// TIA Portal V21 export
// export: Created 2026-11-10T19:11:42.2574666Z, ExportSetting WithDefaults, DisplayName Totally Integrated Automation Portal, DisplayVersion V21 Update 3, DisplayName STEP 7 Professional, DisplayVersion V21 Update 3, DisplayName STEP 7 Safety, DisplayVersion V21, DisplayName Tech WebApplication, DisplayVersion V21, DisplayName WinCC Basic/Comfort/Advanced, DisplayVersion V21 Update 3, DisplayName WinCC Unified, DisplayVersion V21 Update 3
DATA_BLOCK "DB_BSEND_SFB"   // DB54
// stored: AutoNumber true, DBAccessibleFromOPCUA true, DBAccessibleFromWebserver true, InstanceOfName BSEND_SFB, OfSystemLibElement BSEND, OfSystemLibVersion 1.2
"BSEND_SFB"
   // VAR_INPUT
   //    REQ : Bool;
   //    R : Bool;
   //    ID : CONN_PRG;
   //    R_ID : CONN_R_ID;
   // END_VAR
   // VAR_OUTPUT
   //    DONE : Bool;
   //    ERROR : Bool;
   //    STATUS : Word;
   // END_VAR
   // VAR_IN_OUT
   //    SD_1 : Variant;
   //    LEN : Word;
   // END_VAR
   // VAR
   //    INDEX : Word;
   // END_VAR
BEGIN
END_DATA_BLOCK
